Staubli VAL3: copyPoint3.pgx

public program copyPoint3(string x_sKey, num x_nTarget, num x_nSource)
  local num l_i
begin
  trajTemp:tTrajItem[x_sKey].pPointItem[x_nTarget].pPointRx=trajTemp:tTrajItem[x_sKey].pPointItem[x_nSource].pPointRx
  //trajTemp:tTrajItem[x_sKey].pPointItem[x_nTarget].pPointRx[1]=trajTemp:tTrajItem[x_sKey].pPointItem[x_nSource].pPointRx[1]
  trajTemp:tTrajItem[x_sKey].pPointItem[x_nTarget].jJointRx=trajTemp:tTrajItem[x_sKey].pPointItem[x_nSource].jJointRx
  trajTemp:tTrajItem[x_sKey].pPointItem[x_nTarget].sID=trajTemp:tTrajItem[x_sKey].pPointItem[x_nSource].sID
  trajTemp:tTrajItem[x_sKey].pPointItem[x_nTarget].bMarked=trajTemp:tTrajItem[x_sKey].pPointItem[x_nSource].bMarked
  trajTemp:tTrajItem[x_sKey].pPointItem[x_nTarget].pInter=trajTemp:tTrajItem[x_sKey].pPointItem[x_nSource].pInter
  trajTemp:tTrajItem[x_sKey].pPointItem[x_nTarget].pParaItem.mMdesc=trajTemp:tTrajItem[x_sKey].pPointItem[x_nSource].pParaItem.mMdesc
  trajTemp:tTrajItem[x_sKey].pPointItem[x_nTarget].pParaItem.nMoveType=trajTemp:tTrajItem[x_sKey].pPointItem[x_nSource].pParaItem.nMoveType
  trajTemp:tTrajItem[x_sKey].pPointItem[x_nTarget].pParaItem.nActionIndex=trajTemp:tTrajItem[x_sKey].pPointItem[x_nSource].pParaItem.nActionIndex
  trajTemp:tTrajItem[x_sKey].pPointItem[x_nTarget].pParaItem.nPercentage=trajTemp:tTrajItem[x_sKey].pPointItem[x_nSource].pParaItem.nPercentage
  trajTemp:tTrajItem[x_sKey].pPointItem[x_nTarget].pParaItem.nDelay=trajTemp:tTrajItem[x_sKey].pPointItem[x_nSource].pParaItem.nDelay
  trajTemp:tTrajItem[x_sKey].pPointItem[x_nTarget].pParaItem.nSigValue=trajTemp:tTrajItem[x_sKey].pPointItem[x_nSource].pParaItem.nSigValue
  trajTemp:tTrajItem[x_sKey].pPointItem[x_nTarget].pParaItem.bSafePoint=trajTemp:tTrajItem[x_sKey].pPointItem[x_nSource].pParaItem.bSafePoint
  for l_i = 0 to 2
    trajTemp:tTrajItem[x_sKey].pPointItem[x_nTarget].pParaItem.iIfItem.nSigType[l_i]=trajTemp:tTrajItem[x_sKey].pPointItem[x_nSource].pParaItem.iIfItem.nSigType[l_i]
    trajTemp:tTrajItem[x_sKey].pPointItem[x_nTarget].pParaItem.iIfItem.nSigIndex[l_i]=trajTemp:tTrajItem[x_sKey].pPointItem[x_nSource].pParaItem.iIfItem.nSigIndex[l_i]
    trajTemp:tTrajItem[x_sKey].pPointItem[x_nTarget].pParaItem.iIfItem.nValue[l_i]=trajTemp:tTrajItem[x_sKey].pPointItem[x_nSource].pParaItem.iIfItem.nValue[l_i]
  endFor
  trajTemp:tTrajItem[x_sKey].pPointItem[x_nTarget].pParaItem.iIfItem.bANDOR[0]=trajTemp:tTrajItem[x_sKey].pPointItem[x_nSource].pParaItem.iIfItem.bANDOR[0]
  trajTemp:tTrajItem[x_sKey].pPointItem[x_nTarget].pParaItem.iIfItem.bANDOR[1]=trajTemp:tTrajItem[x_sKey].pPointItem[x_nSource].pParaItem.iIfItem.bANDOR[1]

end
